(* IEC 61131-3 sources: plc-st-coding-agent/progress/evidence/f14_v9_temperature_minimal_20261113/native_compile_evidence, 1 file *)

(* ---- candidate.st ---- *)
FUNCTION_BLOCK FB_TemperatureControl
VAR_INPUT
    TemperatureSensorInput : REAL;
    SetTemperature : REAL;
END_VAR
VAR_OUTPUT
    CurrentTemperature : REAL;
    SetTempDisplay : REAL;
    HeaterStatus : BOOL;
    OverheatProtection : BOOL;
    HeaterOutput : BOOL;
END_VAR
VAR
    sensor_fault : BOOL;
    heater_request : BOOL;
    overheat_active : BOOL;
    tmp_heater_in : BOOL;
    HeatingTimer : TON;
    CoolingTimer : TON;
END_VAR

(* ENGINEERING_CONTRACT
   O1 CurrentTemperature: always copies TemperatureSensorInput; no fault suppression; units = input units (PUB006/PUB007).
   O2 SetTempDisplay: always copies SetTemperature; units same as input (PUB006/PUB007).
   O3 HeaterStatus: copies final HeaterOutput; true while actual heater command active (PUB006/PUB007).
   O4 OverheatProtection: latched TRUE when HeatingTimer reaches strictly more than T#5S; holds TRUE while CoolingTimer < T#3S; auto-clears after T#3S; no external reset (PUB005/PUB006).
   O5 HeaterOutput: TRUE when sensor input in [0,100] and TemperatureSensorInput < SetTemperature and not overheat-active; FALSE on sensor fault, overheat, or temp >= set (PUB003/PUB004/PUB005/PUB008).
   State retention: OverheatProtection retained during 3s wait; HeatingTimer resets whenever HeaterOutput is false; CoolingTimer resets when overheat inactive.
   Same-scan priority: overheat set and HeaterOutput forced FALSE in same timer-trigger scan; when cooling timer completes, HeaterOutput may turn on same scan if setpoint condition still true.
   Boundaries: strict < for low-temperature start; fault uses <0.0 or >100.0; exact 0/100 valid; overheat threshold uses T#5S1MS to satisfy strict > T#5S; cooldown threshold T#3S uses >=.
*)
(* CONTRACT_RULES [] *)

sensor_fault := (TemperatureSensorInput < 0.0) OR (TemperatureSensorInput > 100.0);
heater_request := (NOT sensor_fault) AND (TemperatureSensorInput < SetTemperature);

(* Desired heating timer enable before possible cooling-timer completion. *)
tmp_heater_in := heater_request AND NOT overheat_active;

(* Strict overheat threshold: T#5S1MS triggers only after more than 5 seconds. *)
HeatingTimer(IN := tmp_heater_in, PT := T#5S1MS);
IF HeatingTimer.Q THEN
    overheat_active := TRUE;
    tmp_heater_in := FALSE;
END_IF;

(* Cooling timer: cooldown exactly T#3S before protection is lifted. *)
CoolingTimer(IN := overheat_active, PT := T#3S);
IF overheat_active AND CoolingTimer.Q THEN
    overheat_active := FALSE;
END_IF;

HeaterOutput := heater_request AND NOT overheat_active;

(* Ensure HeatingTimer starts immediately when heater turns on in this scan.
   Also reset immediately when heater turns off to avoid one-scan timer drift. *)
IF HeaterOutput AND NOT tmp_heater_in THEN
    HeatingTimer(IN := TRUE, PT := T#5S1MS);
ELSIF (NOT HeaterOutput) AND tmp_heater_in THEN
    HeatingTimer(IN := FALSE, PT := T#5S1MS);
END_IF;

CurrentTemperature := TemperatureSensorInput;
SetTempDisplay := SetTemperature;
HeaterStatus := HeaterOutput;
OverheatProtection := overheat_active;

END_FUNCTION_BLOCK
